// TIA Portal V21 export
// export: Created 2026-11-08T21:35:29.8520864Z, ExportSetting WithDefaults, DisplayName Totally Integrated Automation Portal, DisplayVersion V21 Update 3, DisplayName STEP 7 Professional, DisplayVersion V21 Update 3, DisplayName STEP 7 Safety, DisplayVersion V21, DisplayName Tech WebApplication, DisplayVersion V21, DisplayName WinCC Basic/Comfort/Advanced, DisplayVersion V21 Update 3, DisplayName WinCC Unified, DisplayVersion V21 Update 3
FUNCTION_BLOCK "FB_StlC_029"   // FB87, STL
TITLE = STL call MOVE_BLK_VARIANT
{ S7_Optimized_Access := 'TRUE' }
VERSION : 0.1
// stored: AutoNumber true, IsRetainMemResEnabled false, MemoryReserve 100, UDAEnableTagReadback false
   VAR_INPUT
      cnt : UDInt;
      si : DInt;
      di : DInt;
   END_VAR
   VAR_OUTPUT
      io : Int;
   END_VAR
   VAR_IN_OUT
      src : Variant;
      dst : Variant;
   END_VAR
BEGIN

NETWORK
TITLE = 029 MOVE_BLK_VARIANT
      CALL  MOVE_BLK_VARIANT
      ( SRC        := #src,
        COUNT      := #cnt,
        SRC_INDEX  := #si,
        DEST_INDEX := #di,
        Ret_Val    := #io,
        DEST       := #dst
      );
END_FUNCTION_BLOCK
